// TIA Portal V21 export
// export: Created 2000-01-01T00:00:00.0000000Z, ExportSetting None
TYPE "UDT_HMI_FIO_BufferConveyor"
   STRUCT
      bManualMode { ExternalWritable := 'False'} : Bool;   // TRUE手动, FALSE自动
      bStartCmd { ExternalWritable := 'False'} : Bool;   // HMI启动命令
      bStopCmd { ExternalWritable := 'False'} : Bool;   // HMI停止命令
      bResetCmd { ExternalWritable := 'False'} : Bool;   // HMI复位命令
      bManualConv1 { ExternalWritable := 'False'} : Bool;   // 手动驱动1号缓冲带
      bManualConv2 { ExternalWritable := 'False'} : Bool;   // 手动驱动2号缓冲带
      bManualConv3 { ExternalWritable := 'False'} : Bool;   // 手动驱动3号缓冲带
      tJamTimeout { ExternalWritable := 'False'} : Time;   // 光电长遮挡卡料超时阈值（默认 T#6s）
      iOccupiedZones { ExternalWritable := 'False'} : Int;   // 状态反馈：当前被占用的缓冲区段数 (0..3)
      bBufferFull { ExternalWritable := 'False'} : Bool;   // 状态反馈：三级缓冲全满标志
      bJamFault { ExternalWritable := 'False'} : Bool;   // 状态反馈：传送带卡料报警
      wStatus { ExternalWritable := 'False'} : Word;   // 状态码：16#0000正常, 16#7000停机, 16#8401卡料超时, 16#8402急停触发
   END_STRUCT;
END_TYPE
